// SIMATIC STEP 7 (V5.x) project EX8
// CPU: CPU 314
// station: Matériel
// station: SIMATIC 300(1)
// station: P_ADR_BUS
// program: Programme S7(1)

ORGANIZATION_BLOCK OB 1
TITLE = "Main Program Sweep (Cycle)"
VERSION : 0.1
VAR_TEMP
  OB1_EV_CLASS : BYTE ;	//Bits 0-3 = 1 (Coming event), Bits 4-7 = 1 (Event class 1)
  OB1_SCAN_1 : BYTE ;	//1 (Cold restart scan 1 of OB 1), 3 (Scan 2-n of OB 1)
  OB1_PRIORITY : BYTE ;	//Priority of OB Execution
  OB1_OB_NUMBR : BYTE ;	//1 (Organization block 1, OB1)
  OB1_RESERVED_1 : BYTE ;	//Reserved for system
  OB1_RESERVED_2 : BYTE ;	//Reserved for system
  OB1_PREV_CYCLE : INT ;	//Cycle time of previous OB1 scan (milliseconds)
  OB1_MIN_CYCLE : INT ;	//Minimum cycle time of OB1 (milliseconds)
  OB1_MAX_CYCLE : INT ;	//Maximum cycle time of OB1 (milliseconds)
  OB1_DATE_TIME : DATE_AND_TIME ;	//Date and time OB1 started
END_VAR
BEGIN
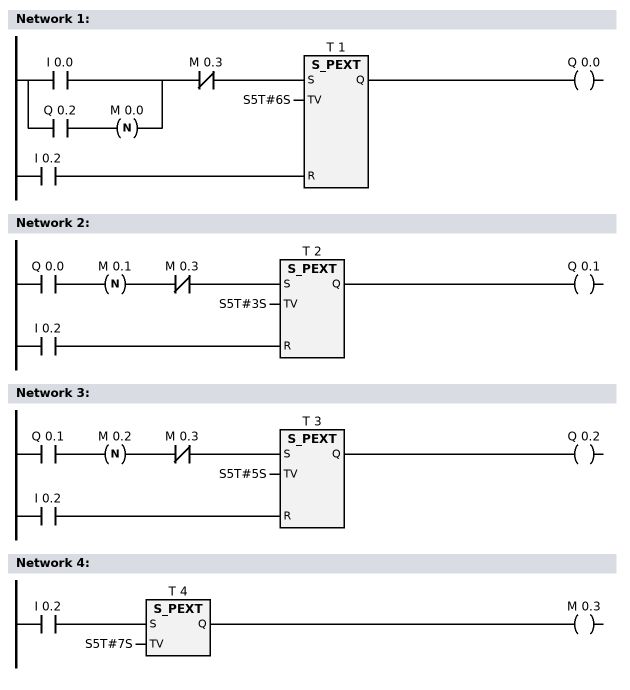
NETWORK
TITLE =
      A(;
      O     I 0.0;
      O(;
      A     Q 0.2;
      FN    M 0.0;
      );
      );
      AN    M 0.3;
      L     S5T#6S;
      SE    T 1;
      A     I 0.2;
      R     T 1;
      NOP   0;
      NOP   0;
      A     T 1;
      =     Q 0.0;
NETWORK
TITLE =
      A     Q 0.0;
      FN    M 0.1;
      AN    M 0.3;
      L     S5T#3S;
      SE    T 2;
      A     I 0.2;
      R     T 2;
      NOP   0;
      NOP   0;
      A     T 2;
      =     Q 0.1;
NETWORK
TITLE =
      A     Q 0.1;
      FN    M 0.2;
      AN    M 0.3;
      L     S5T#5S;
      SE    T 3;
      A     I 0.2;
      R     T 3;
      NOP   0;
      NOP   0;
      A     T 3;
      =     Q 0.2;
NETWORK
TITLE =
      A     I 0.2;
      L     S5T#7S;
      SE    T 4;
      NOP   0;
      NOP   0;
      NOP   0;
      A     T 4;
      =     M 0.3;
END_ORGANIZATION_BLOCK
